(* CODESYS project i_camera.library
   DefaultNamespace: KOSTAL.AF2024.Drivers.Camera.I_Camera
   DocFormat: reStructuredText
   Description: Base Interface for Camera Systems
   Author: Frank Dümpelmann / Martin Hundt
   Title: KOSTAL.AF2024.Drivers.Camera.I_Camera
   Version: 2.0.0.0
   Company: KOSTAL GmbH & Co.KG
   Placeholder: KOSTAL.AF2024.Drivers.Camera.I_Camera

Project tree, tasks and I/O mapping:
  libraries: KOSTAL.AF2024.Core.Process, 1.0.0.0 (KOSTAL GmbH & Co.KG); KOSTAL.AF2024.Core.Settings, 1.0.0.0 (KOSTAL GmbH & Co.KG); KOSTAL.AF2024.Core.System, 1.0.0.0 (KOSTAL GmbH & Co.KG)
  Project Information/
    function F_GetCompany [ST]
    function F_GetTitle [ST]
    function F_GetVersion [ST]
  Version/
    global variables Global_Version
  interface I_Camera: Ex_SetProgramNumber, Ex_Trigger, Ex_Trigger_ProgramNumber, ResultPass, State
  interface I_CameraWithFeedback: ProgramNumber
*)

// Version/Global_Version
{attribute 'TcGenerated'}
{attribute 'no-analysis'}
{attribute 'linkalways'}
// This function has been automatically generated from the project information.
VAR_GLOBAL CONSTANT
	{attribute 'const_non_replaced'}
	stLibVersion_KOSTAL_AF2024_Drivers_Camera_I_Camera : ST_LibVersion := (iMajor := 2, iMinor := 0, iBuild := 0, iRevision := 0, nFlags := 0, sVersion := '2.0.0.0');
END_VAR

// Project Information/F_GetCompany
// This function has been automatically generated from the project information.
{attribute 'signature_flag' := '1073741824'}
{attribute 'TcGenerated'}
{attribute 'no-analysis'}
FUNCTION F_GetCompany : WSTRING
VAR_INPUT
	
END_VAR

F_GetCompany := "KOSTAL GmbH & Co.KG";

END_FUNCTION

// Project Information/F_GetTitle
// This function has been automatically generated from the project information.
{attribute 'signature_flag' := '1073741824'}
{attribute 'TcGenerated'}
{attribute 'no-analysis'}
FUNCTION F_GetTitle : WSTRING
VAR_INPUT
	
END_VAR

F_GetTitle := "KOSTAL.AF2024.Drivers.Camera.I_Camera";

END_FUNCTION

// I_Camera
INTERFACE I_Camera EXTENDS KOSTAL_AF2024_Core_System.I_Interface

METHOD PUBLIC Ex_SetProgramNumber	:	BOOL
VAR_INPUT
	ProgramNumber	: UINT;
END_VAR
END_METHOD

METHOD PUBLIC Ex_Trigger	:	BOOL
END_METHOD

METHOD PUBLIC Ex_Trigger_ProgramNumber	:	BOOL
VAR_INPUT
	ProgramNumber	: UINT;
END_VAR
END_METHOD

PROPERTY ResultPass : BOOL
GET
END_GET
END_PROPERTY

PROPERTY PUBLIC State : KOSTAL_AF2024_Core_Process.I_T_plcState
GET
END_GET
END_PROPERTY

END_INTERFACE

// Project Information/F_GetVersion
// This function has been automatically generated from the project information.
{attribute 'signature_flag' := '1073741824'}
{attribute 'TcGenerated'}
{attribute 'no-analysis'}
FUNCTION F_GetVersion : ST_LibVersion
VAR_INPUT
	
END_VAR

F_GetVersion.iMajor := 2;
F_GetVersion.iMinor := 0;
F_GetVersion.iBuild := 0;
F_GetVersion.iRevision := 0;
F_GetVersion.sVersion := '2.0.0.0';
F_GetVersion.nFlags := 0;

END_FUNCTION

// I_CameraWithFeedback
INTERFACE I_CameraWithFeedback EXTENDS I_Camera

PROPERTY ProgramNumber : UINT
GET
END_GET
END_PROPERTY

END_INTERFACE
